SUBAPPLICATION AX_TO_BG_PUBLISH (* Fertiger AX-Zustand auf Hintergrundfarbe (SoftKey+AUX, GreenWhiteBackground3_AXC) + lokalen State-Publish - wie AX_TO_QXA_BG_PUBLISH, aber ohne physischen Ausgang. INIT per Auto-Verteilung. *)
  (* Standard: 61499-2; Description: Copyright (c) 2026 Meisterschulen am Ostbahnhof This program and the accompanying materials are made available under the terms of the Eclipse Public License 2.0 which is available at https://www.eclipse.org/legal/epl-2.0/ SPDX-License-Identifier: EPL-2.0 *)
  (* Version 1.0, 2026-10-17, Franz Höpfinger, Meisterschulen am Ostbahnhof, initial implementation - AX_SPLIT_2 + GreenWhiteBackground3_AXC + AX_PUBLISH_1 aus Baender_EinAus.SUB (Background_Alle/AX_PUBLISH_Alle) als wiederverwendbarer Baustein. *)
  PACKAGE MyLib::sys;
  IMPORT isobus::UT::Q::const::IDs::ID_NULL;
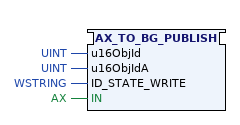
  VAR_INPUT
    u16ObjId : UINT := ID_NULL; (* Object ID Softkey - traegt die Hintergrundfarbe *)
    u16ObjIdA : UINT := ID_NULL; (* Object ID AuxFunction2 (Joystick) - zeigt Hintergrundfarbe am Aux-Handle mit *)
    ID_STATE_WRITE : WSTRING; (* Lokale Publish-Adresse (ACTION=WRITE) fuer den Zustand - wird remote abonniert *)
  END_VAR
  SOCKETS
    IN : adapter::types::unidirectional::AX; (* Fertiger AX-Zustand - wird auf Hintergrund+Publish verteilt *)
  END_SOCKETS
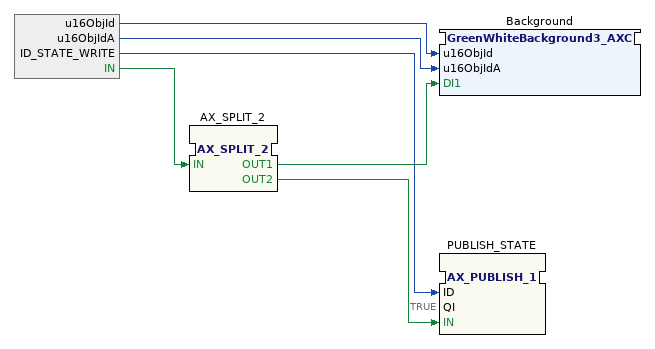
  FBS
    AX_SPLIT_2 : adapter::events::unidirectional::AX_SPLIT_2; (* Adapter-Fanout ist strikt 1:1 *)
    PUBLISH_STATE : adapter::net::AX_PUBLISH_1(QI := TRUE);
  END_FBS
  SUBAPPS
    Background : MyLib::sys::GreenWhiteBackground3_AXC;
  END_SUBAPPS
  DATA_CONNECTIONS
    u16ObjId TO Background.u16ObjId;
    u16ObjIdA TO Background.u16ObjIdA;
    ID_STATE_WRITE TO PUBLISH_STATE.ID;
  END_CONNECTIONS
  ADAPTER_CONNECTIONS
    IN TO AX_SPLIT_2.IN;
    AX_SPLIT_2.OUT1 TO Background.DI1;
    AX_SPLIT_2.OUT2 TO PUBLISH_STATE.IN;
  END_CONNECTIONS
END_SUBAPPLICATION
